Universal Robots PolyScope program: ConfProg.urp

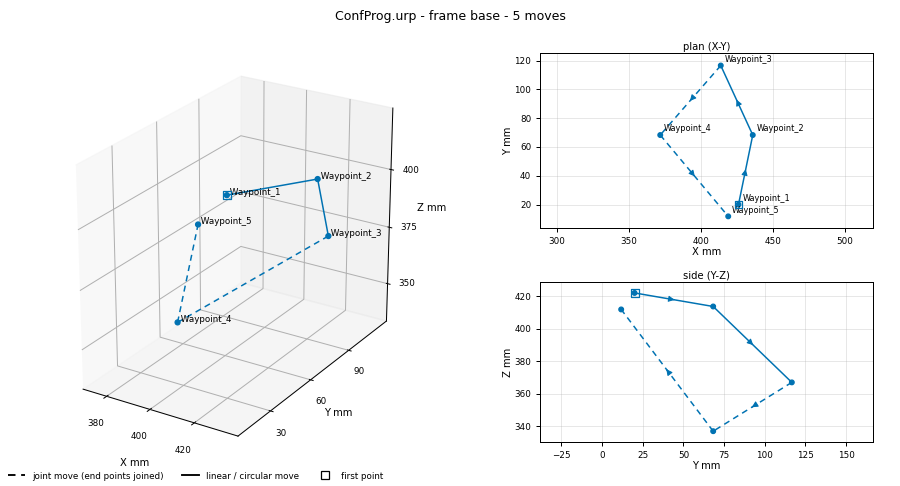
[picture p0: tool path of ConfProg.urp in frame base, 5 of 5 moves have a stored position in this frame; points joined in program order, loops and branches not executed]
Program ConfProg (createdIn=3.0.0 lastSavedIn=3.0.0 directory=/programs installation=default)
Robot Program (runOnlyOnce=true motionType=MoveJ speed=1.047198 acceleration=1.396263 useActiveTCP=false)
  'Program generated by RoboDK v6.0.7 for ABB IRB 120-3/0.6 on XX/XX/XXXX 18:00:00'
  'Using nominal kinematics.'
  'Using Ref. Frame S: p[1.234570, -0.098765, 0.050500, 0.000000, 0.000000, 0.523599]'
  'Using TCP Tool S: p[0.010000, 0.020000, 0.150000, 0.000000, 0.000000, 0.000000]'
  Script: set_tcp(p[0.010000, 0.020000, 0.150000, 0.000000, 0.000000, 0.000000])
  MoveL speed 250 mm/s, acceleration 1200 mm/s^2 (useActiveTCP=true)
    Waypoint Waypoint_1: TCP in base x=426.318 y=20 z=422.034 mm, rx=0.1383 ry=2.2532 rz=-0.2966 rad; joints [0, -10, 20, 0, 30, 0] deg; flange x=317.789 y=39.504 z=526.155 mm, rx=0.1383 ry=2.2532 rz=-0.2966 rad
    Waypoint Waypoint_2: TCP in base x=436.232 y=68.297 z=413.715 mm, rx=0.1383 ry=2.2532 rz=-0.2966 rad; joints [185, -10, 20, 190, 30, -270] deg; flange x=327.703 y=87.801 z=517.836 mm, rx=0.1383 ry=2.2532 rz=-0.2966 rad
    Waypoint Waypoint_3: TCP in base x=414.005 y=116.593 z=367.095 mm, rx=0.1383 ry=2.2532 rz=-0.2966 rad; joints [-185, -60, 100, -190, -30, 370] deg; flange x=305.476 y=136.097 z=471.216 mm, rx=0.1383 ry=2.2532 rz=-0.2966 rad
  Script: movej([0.174533, 0.349066, -0.523599, 0.698132, -0.872665, 1.047198],1.20000,0.75000,0,0.0000)
  MoveJ speed 42.97 deg/s, acceleration 68.75 deg/s^2 (useActiveTCP=true)
    Waypoint Waypoint_4: TCP in base x=371.953 y=68.296 z=337.111 mm, rx=0.1383 ry=2.2532 rz=-0.2966 rad; joints [10, 20, -30, 40, -50, 60] deg; flange x=263.425 y=87.801 z=441.232 mm, rx=0.1383 ry=2.2532 rz=-0.2966 rad
  Script: movej([-2.967060, 0.785398, -0.785398, -2.967060, 1.570796, -3.124139],1.20000,0.75000,0,0.0000)
  MoveJ speed 42.97 deg/s, acceleration 68.75 deg/s^2 (useActiveTCP=true)
    Waypoint Waypoint_5: TCP in base x=419.189 y=11.793 z=411.899 mm, rx=0.1383 ry=2.2532 rz=-0.2966 rad; joints [-170, 45, -45, -170, 90, -179] deg; flange x=310.661 y=31.298 z=516.02 mm, rx=0.1383 ry=2.2532 rz=-0.2966 rad
  'Circular move (R405.1 mm)'
  Script: movec(p[0.973908, -0.353337, 0.382202, -0.503745, 2.359457, 0.000119],p[0.408367, 0.083800, 0.505120, -0.487372, 1.445847, -0.747268],1.20000,0.25000,0.0000)
